(* IEC 61131-3 sources: 89152_FlorisHendrix_AfstudeerProject/89152_FlorisHendrix_ExamenProject/Stations/MachineControl/MachineControl/Network/KTS_Network, 1 file *)

(* ---- ONE_KTS_Network_Table.st ---- *)
#define OBJECTS_CONFIG

//Define part of class HWKVarSizeFIFO
#define _HWKBUF_MEMID 16#1E3B0000
//Define part of class SdiasBase
//Address to access the Dataobject list via SPI SDO Read
#define SDIAS_SPI_DATA_OBJECT_LIST_PAGE_ADDRESS               16#FFFF
#define SDIAS_SPI_DATA_OBJECT_LIST_PAGE_OFFSET                16#00
#define SDIAS_SPI_DATA_OBJECT_LIST_IDENTIFIER                 16#12345678

//Defines the number of optional list elements in the SPI List

#define SDIAS_SPI_NUMBER_OF_OPTIONAL_ELEMENTS                 16

#define SDIAS_SPI_HEADER_BEFORE_OPTIONAL_ELEMENTS             16#18
#define SDIAS_SPI_HARDWARE_VERSION_OFFSET                     16#C
#define SDIAS_SPI_VENDOR_ID_OFFSET                            16#0

#define SDIAS_SPI_MASTER_ADRESS_TRANSMIT_BUFFER0              16#0000
#define SDIAS_SPI_MASTER_ADRESS_TRANSMIT_BUFFER1              16#0080
#define SDIAS_SPI_MASTER_ADRESS_RECEIVE_BUFFER0               16#0000
#define SDIAS_SPI_MASTER_ADRESS_RECEIVE_BUFFER1               16#0080
#define SDIAS_SPI_MASTER_ADRESS_PAGE_ADRESS                   16#0100
#define SDIAS_SPI_MASTER_ADRESS_PREDEFINED_COMMAND_REGISTER   16#0102
#define SDIAS_SPI_MASTER_ADRESS_SINGLE_COMMAND_REGISTER       16#0103
#define SDIAS_SPI_MASTER_ADRESS_STATUS_REGISTER               16#0104
#define SDIAS_SPI_MASTER_ADRESS_REQUEST_REGISTER              16#0105
#define SDIAS_SPI_MASTER_ADRESS_GRANT_REGISTER                16#0106
#define SDIAS_SPI_MASTER_ADRESS_CLEAR_REQUEST_REGISTER        16#0107
#define SDIAS_SPI_MASTER_ADRESS_FEATURE_REGISTER              16#0108

#define SDIAS_SPI_MASTER_SOFTWARE_REQUEST                     1

#define SDIAS_SPI_MASTER_COMMAND_PAGE_READ                    16#01
#define SDIAS_SPI_MASTER_COMMAND_PAGE_PROGRAM                 16#02
#define SDIAS_SPI_MASTER_COMMAND_SECTOR_ERASE                 16#03
#define SDIAS_SPI_MASTER_COMMAND_REBOOT_FPGA                  16#F0

#define SDIAS_SPI_MASTER_STATE_BUSY                           16#00
#define SDIAS_SPI_MASTER_STATE_READY                          16#01

#define SDIAS_SPI_SECTOR_SIZE                                 65536 // 256*256
#define SDIAS_SPI_PAGE_SIZE                                   256

#define SDIAS_SPI_WRITE_MAX_RETRIES                           2
#define SDIAS_SPI_TIMEOUT                                     500  //timeout for spi accesses
#define SDIAS_SPI_LOCK_TIMEOUT                                6   //this value is multiplied with the buscycletime [µs] (6*1000=6.000 msec timeout)

//SPI List IDs
#define SDIAS_SPI_IDENTIFICATION_LIST_ID  1
#define SDIAS_SPI_FLASH_CONFIGURATION_ID  2
#define SDIAS_SPI_VENDOR_NAME_ID          3
#define SDIAS_SPI_DEVICE_NAME_ID          4
#define SDIAS_SPI_SERIAL_NUMBER_ID        5
#define SDIAS_SPI_ORDERING_NUMBER_ID      6
#define SDIAS_SPI_DOCUMENTATION_PDF_ID    7
#define SDIAS_SPI_CALIB_DATA_ID           10
#define SDIAS_SPI_PDO_INFORMATION_ID      128

//SPI Access
#define SDIAS_SPI_ACCESS_ID_HW_TREE          1
#define SDIAS_SPI_ACCESS_ID_HWK_INTERNAL     2
#include "..\..\Class\SdiasManager\SdiasManager.h"
#include "..\..\Class\SdiasBase\SdiasBase.h"
#include "..\..\Class\HwControl\HwControl.h"
#include "..\..\Source\interfaces\lsl_st_hardwaretree.h"
#include "..\..\Source\interfaces\lsl_st_mt.h"
//Define part of class SdiasSDCIMaster
#define SSDCIM_SDO_LOCK    16#1B3D5F2A
#define SSDCIM_SDO_UNLOCK  16#2E9A3C57
#include "..\..\Source\BusInterface.h"
#include "..\..\Class\SdiasSDCIMaster\SdiasSDCIMaster.h"
//Define part of class IIO041
#define IIO041_DEVICE_ID  1077
#include "..\..\Class\KTS_TimeStamp\KTS_TimeStamp_SDCI_Parameters.h"
#include <.\lsl_st_mt.h>

FUNCTION GLOBAL TAB ONE_KTS_Network
-1$UINT, 0$UINT,
0$UINT, 0$UINT,

16$UDINT,
TO_UDINT(794617671), "CriticalSection", 0$UINT, 4$UINT, 1$UINT,
TO_UDINT(2647432661), "HWKVarSizeFIFO", 1$UINT, 0$UINT, 1$UINT,
TO_UDINT(3248397833), "IIO041", 1$UINT, 17$UINT, 1$UINT,
TO_UDINT(2039520762), "KTS_Read", 0$UINT, 0$UINT, 1$UINT,
TO_UDINT(3289613158), "KTS_TimeStamp", 0$UINT, 0$UINT, 1$UINT,
TO_UDINT(2225119864), "MerkerEx", 1$UINT, 22$UINT, 1$UINT,
TO_UDINT(933570811), "RAMex", 1$UINT, 17$UINT, 2$UINT,
TO_UDINT(205726265), "SDCIDevice", 1$UINT, 9$UINT, 0$UINT,
TO_UDINT(1321842971), "SDCIDevice_AsyncPara", 1$UINT, 4$UINT, 1$UINT,
TO_UDINT(2258655160), "SDCIPort", 1$UINT, 0$UINT, 4$UINT,
TO_UDINT(3175101883), "SdiasBase", 1$UINT, 60$UINT, 0$UINT,
TO_UDINT(2874110376), "SdiasSDCIMaster", 1$UINT, 15$UINT, 0$UINT,
TO_UDINT(1850111279), "String", 1$UINT, 11$UINT, 1$UINT,
TO_UDINT(2898603620), "StringInternal", 1$UINT, 85$UINT, 0$UINT,
TO_UDINT(2408581120), "StringRAM", 1$UINT, 10$UINT, 2$UINT,
TO_UDINT(3232495061), "VirtualBaseInit", 1$UINT, 3$UINT, 0$UINT,

1$UINT, TO_UDINT(2270667760), "IIO0411\_BASE\PDOPROTECTION",

1$UINT, TO_UDINT(3344372028), "IIO0411\_BASE\HWKVARSIZEFIFO1",

_NO_ATTR, TO_UDINT(4207004045), "IIO0411",

_NO_ATTR, TO_UDINT(2039520762), "KTS_READ",

_NO_ATTR, TO_UDINT(667498585), "KTS_TIMESTAMP1",

1$UINT, TO_UDINT(1001843434), "IIO0411\_BASE\_BASE\SERIALNOSTR\MERKEREX0",

1$UINT, TO_UDINT(524577153), "KTS_READ\STRINGPRODUCTNAME\DATABUFFER",
1$UINT, TO_UDINT(558793340), "KTS_READ\STRINGVENDORNAME\DATABUFFER",

_NO_ATTR, TO_UDINT(729601649), "SDCIDEVICE_ASYNCPARA_KTS_TIMESTAMP",

1$UINT, TO_UDINT(2446752732), "IIO0411\SDCIPORT1",
1$UINT, TO_UDINT(148843110), "IIO0411\SDCIPORT2",
1$UINT, TO_UDINT(2144869104), "IIO0411\SDCIPORT3",
1$UINT, TO_UDINT(3787231059), "IIO0411\SDCIPORT4",

1$UINT, TO_UDINT(2058560523), "IIO0411\_BASE\_BASE\SERIALNOSTR",

1$UINT, TO_UDINT(901476136), "KTS_READ\STRINGPRODUCTNAME",
1$UINT, TO_UDINT(1642288413), "KTS_READ\STRINGVENDORNAME",

//Internal connections
0$UDINT,
12$UDINT,
TO_UDINT(2), "SerialNoStr", TO_UDINT(13),
TO_UDINT(2), "PdoProtection", TO_UDINT(0),
TO_UDINT(2), "HWKVarSizeFIFO1", TO_UDINT(1),
TO_UDINT(2), "SDCIPort1", TO_UDINT(9),
TO_UDINT(2), "SDCIPort2", TO_UDINT(10),
TO_UDINT(2), "SDCIPort3", TO_UDINT(11),
TO_UDINT(2), "SDCIPort4", TO_UDINT(12),
TO_UDINT(3), "StringVendorName", TO_UDINT(15),
TO_UDINT(3), "StringProductName", TO_UDINT(14),
TO_UDINT(13), "MerkerEx0", TO_UDINT(5),
TO_UDINT(14), "DataBuffer", TO_UDINT(6),
TO_UDINT(15), "DataBuffer", TO_UDINT(7),
0$UDINT,
11$UDINT,
TO_UDINT(3), "SDCI_Device", TO_UDINT(4), "ClassState",
TO_UDINT(3), "SDCI_Device_Async", TO_UDINT(8), "CmdState",
TO_UDINT(4), "SdciIn", TO_UDINT(9), "ClassSvr",
TO_UDINT(8), "ToDevice", TO_UDINT(4), "ClassState",
TO_UDINT(9), "ToMaster", TO_UDINT(2), "ClassState",
TO_UDINT(10), "ToMaster", TO_UDINT(2), "ClassState",
TO_UDINT(11), "ToMaster", TO_UDINT(2), "ClassState",
TO_UDINT(12), "ToMaster", TO_UDINT(2), "ClassState",
TO_UDINT(13), "DataBuffer", TO_UDINT(5), "m_udLength",
TO_UDINT(14), "DataBuffer", TO_UDINT(6), "m_udLength",
TO_UDINT(15), "DataBuffer", TO_UDINT(7), "m_udLength",

//Initialization values
0$UDINT,
28$UDINT,
TO_UDINT(1), "MaxBufferSize", TO_UDINT(1024),//|KTS_Network._base\IIO0411\HWKVarSizeFIFO1.MaxBufferSize;
TO_UDINT(2), "LEDControl", TO_UDINT(0),//|KTS_Network.IIO0411.LEDControl;
TO_UDINT(2), "Place", TO_UDINT(2),//|KTS_Network.IIO0411.Place;
TO_UDINT(2), "Required", TO_UDINT(1),//|KTS_Network.IIO0411.Required;
TO_UDINT(2), "StartInInit", TO_UDINT(1),//|KTS_Network.IIO0411.StartInInit;
TO_UDINT(2), "MaxBufferSize", TO_UDINT(1024),//|KTS_Network.IIO0411.MaxBufferSize;
TO_UDINT(2), "WaitTimeReconnect", TO_UDINT(500),//|KTS_Network.IIO0411.WaitTimeReconnect;
TO_UDINT(4), "MinCycleTime", TO_UDINT(0),//|KTS_Network.KTS_TimeStamp1.MinCycleTime;
TO_UDINT(4), "Required", TO_UDINT(0),//|KTS_Network.KTS_TimeStamp1.Required;
TO_UDINT(4), "SkipEndianSwap", TO_UDINT(1),//|KTS_Network.KTS_TimeStamp1.SkipEndianSwap;
TO_UDINT(4), "SkipEndianSwapAsy", TO_UDINT(1),//|KTS_Network.KTS_TimeStamp1.SkipEndianSwapAsy;
TO_UDINT(4), "StartUpMode", TO_UDINT(_SDCI),//|KTS_Network.KTS_TimeStamp1.StartUpMode;
TO_UDINT(4), "ReadPdoSize", TO_UDINT(16),//|KTS_Network.KTS_TimeStamp1.ReadPdoSize;
TO_UDINT(4), "WritePdoSize", TO_UDINT(0),//|KTS_Network.KTS_TimeStamp1.WritePdoSize;
TO_UDINT(4), "AutoConnectTime", TO_UDINT(0),//|KTS_Network.KTS_TimeStamp1.AutoConnectTime;
TO_UDINT(4), "ModeChangeTime", TO_UDINT(500),//|KTS_Network.KTS_TimeStamp1.ModeChangeTime;
TO_UDINT(5), "ThreadSafe", TO_UDINT(0),//|KTS_Network.SerialNoStr\_base\_base\IIO0411\MerkerEx0.ThreadSafe;
TO_UDINT(6), "ThreadSafe", TO_UDINT(0),//|KTS_Network.StringProductName\KTS_Read\DataBuffer.ThreadSafe;
TO_UDINT(7), "ThreadSafe", TO_UDINT(0),//|KTS_Network.StringVendorName\KTS_Read\DataBuffer.ThreadSafe;
TO_UDINT(8), "useBufferedAsyCmds", TO_UDINT(1),//|KTS_Network.SDCIDevice_AsyncPara_KTS_TimeStamp.useBufferedAsyCmds;
TO_UDINT(8), "TimeoutAsyCmd", TO_UDINT(10000),//|KTS_Network.SDCIDevice_AsyncPara_KTS_TimeStamp.TimeoutAsyCmd;
TO_UDINT(9), "PortNo", TO_UDINT(0),//|KTS_Network.IIO0411\SDCIPort1.PortNo;
TO_UDINT(10), "PortNo", TO_UDINT(1),//|KTS_Network.IIO0411\SDCIPort2.PortNo;
TO_UDINT(11), "PortNo", TO_UDINT(2),//|KTS_Network.IIO0411\SDCIPort3.PortNo;
TO_UDINT(12), "PortNo", TO_UDINT(3),//|KTS_Network.IIO0411\SDCIPort4.PortNo;
TO_UDINT(13), "SingleRealloc", TO_UDINT(1),//|KTS_Network._base\_base\IIO0411\SerialNoStr.SingleRealloc;
TO_UDINT(14), "SingleRealloc", TO_UDINT(1),//|KTS_Network.KTS_Read\StringProductName.SingleRealloc;
TO_UDINT(15), "SingleRealloc", TO_UDINT(1),//|KTS_Network.KTS_Read\StringVendorName.SingleRealloc;

//Symbolic initialization values
0$UDINT,
0$UDINT,

//Initialization of string values
0$UDINT,
0$UDINT,

//Configuration of tasks (RealTime, Cyclic, Background)
0$UDINT,
1$UDINT,
TO_UDINT(3), (10)$UDINT, 4194303$DINT, 	//KTS_READ

0$UDINT,
2$UDINT,
TO_UDINT(3), (50)$UDINT, 4194303$DINT, 	//KTS_READ
TO_UDINT(8), (10)$UDINT, 4194303$DINT, 	//SDCIDEVICE_ASYNCPARA_KTS_TIMESTAMP

0$UDINT,
0$UDINT,

//External connections
0$UDINT,
2$UDINT,
TO_UDINT(2), "SdiasIn", C_DIR, TO_UDINT(1007630054), "SdiasPLC1\SdiasHubBase1","ClassSvr",
TO_UDINT(3), "coCSVFile", C_DIR, TO_UDINT(3500464540), "FileBaseCsv1","ClassSvr",

//Magic internal connections
0$UDINT,
3$UDINT,
TO_UDINT(1), "MaxBufferSize", TO_UDINT(2), "MaxBufferSize",
TO_UDINT(6), "UseFile", TO_UDINT(14), "UseFile",
TO_UDINT(7), "UseFile", TO_UDINT(15), "UseFile",

//Configuration of timeslots of tasks (RealTime, Cyclic)
#ifdef __LSLLDR_TIMESLOTS__
0$UDINT,
0$UDINT,

0$UDINT,
0$UDINT,

#endif //__LSLLDR_TIMESLOTS__

//MultiMaster connections
#ifdef __LSLLDR_MULTIMASTER__
0$UDINT,
0$UDINT,
#endif //__LSLLDR_MULTIMASTER__

//Configuration for task ID (RealTime, CyclicTime)
#ifdef __LSLLDR_TASKID__
"\\\\TASKS2  "
0$UDINT,
1$UDINT,
(0)$UDINT, 	//KTS_READ

0$UDINT,
2$UDINT,
(0)$UDINT, 	//KTS_READ
(0)$UDINT, 	//SDCIDEVICE_ASYNCPARA_KTS_TIMESTAMP

0$UDINT,
0$UDINT,

#endif //__LSLLDR_TASKID__

END_FUNCTION
